(*
SPDX-License-Identifier: MIT
License: https://opensource.org/license/mit
*)

(*!
<summary>Owns a nested group of failure scenarios.</summary>
<description>
Owns persistent child storage and fixed parent associations. Use in one task without reentry.
Children is borrowed and must not be modified by application code. Constructor callbacks are not used.
</description>
*)

{attribute 'no_assign'}
{attribute 'no_explicit_call' := 'do not call this function block directly'}
FUNCTION_BLOCK NestedFailureTestGroup EXTENDS TOF_Testing.TestGroup<1>
VAR_STAT
	//! <summary>Class name shared by all instances of this function block.</summary>
	{attribute 'hide'}
	_ClassName : STRING := __POUNAME();
END_VAR
VAR
	{attribute 'hide'}
	{attribute 'init_namespace'}
	_NamespaceName : STRING;
END_VAR
VAR_OUTPUT
	//! <summary>Owned nested failure group.</summary>
	Failures : FailureTestGroup(name := "Failures", parent := THIS^);
END_VAR
VAR
	_Children : ARRAY [0.._ChildCount - 1] OF TOF_Testing.ITestElement :=
	[
		Failures
	];
END_VAR

//! <summary>Borrows the concrete class name for the lifetime of this instance; callers must not modify it.</summary>
{attribute 'monitoring' := 'call'}
PROPERTY ClassName : REFERENCE TO STRING
GET
ClassName REF= _ClassName;
END_GET
END_PROPERTY

//! <summary>Borrows the compiler-initialized namespace; callers must not modify the returned reference.</summary>
{attribute 'monitoring' := 'call'}
PROPERTY NamespaceName : REFERENCE TO STRING
GET
NamespaceName REF= _NamespaceName;
END_GET
END_PROPERTY

//! <summary>Reports the complete concrete instance size, excluding separately allocated storage.</summary>
{attribute 'monitoring' := 'call'}
PROPERTY SelfSize : ULINT
GET
SelfSize := XSIZEOF(THIS^);
END_GET
END_PROPERTY

//! <summary>Borrows the fixed array of this concrete group; do not modify it.</summary>
{attribute 'monitoring' := 'call'}
PROPERTY Children : REFERENCE TO ARRAY [0.._ChildCount - 1] OF TOF_Testing.ITestElement
GET
Children REF= _Children;
END_GET
END_PROPERTY

END_FUNCTION_BLOCK

(* stored: Version 1.1.0.1
   POU NestedFailureTestGroup: Id {2bc23527-1daf-4abd-bed3-caebe4b500c0}, SpecialFunc None
   Property ClassName: Id {c32b4745-93d2-4037-b09c-b2be7b8a77fc}
   Get Get: Id {c5b61716-3ced-4150-abfc-2748164f7755}
   Property NamespaceName: Id {59e89a18-1d31-4762-899a-5a87b553bb1e}
   Get Get: Id {d2d41a5d-6fb9-4f17-818c-38b8ce12f5f3}
   Property SelfSize: Id {e5b6086d-79f7-47a9-b0ad-adb55503580e}
   Get Get: Id {1fcea326-01dc-4456-834e-870bda89647a}
   Property Children: Id {df64e894-f96d-4985-b006-5f3ebcdf6b35}
   Get Get: Id {69ceddb7-4c3f-466b-8134-c5718cdb7044} *)
